// TIA Portal V21 export
// export: Created 2026-11-11T00:47:26.5977342Z, ExportSetting WithDefaults, DisplayName Totally Integrated Automation Portal, DisplayVersion V21 Update 3, DisplayName STEP 7 Professional, DisplayVersion V21 Update 3, DisplayName STEP 7 Safety, DisplayVersion V21, DisplayName Tech WebApplication, DisplayVersion V21, DisplayName WinCC Basic/Comfort/Advanced, DisplayVersion V21 Update 3, DisplayName WinCC Unified, DisplayVersion V21 Update 3
FUNCTION_BLOCK "FB_Fbd_ex103"   // FB115, FBD
{ S7_Optimized_Access := 'TRUE' }
VERSION : 0.1
// stored: AutoNumber true, IsIECCheckEnabled false, IsRetainMemResEnabled false, MemoryReserve 100, SetENOAutomatically false, UDAEnableTagReadback false
   VAR_INPUT
      v_ob_nr : Int;
   END_VAR
   VAR_OUTPUT
      v_cycle : UDInt;
      v_phase : UDInt;
      v_status : Word;
      v_ret_val : Int;
   END_VAR
BEGIN

REGION Network 1: QRY_CINT - Query cyclic interrupt parameters
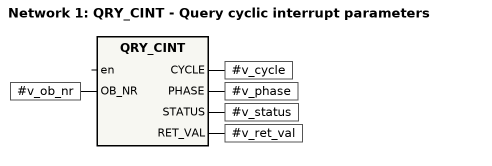
   #v_ret_val := QRY_CINT(OB_NR := #v_ob_nr, CYCLE => #v_cycle, PHASE => #v_phase, STATUS => #v_status);
END_REGION
END_FUNCTION_BLOCK
